Fanuc KAREL source: KD00028.KL

PROGRAM KD00028
%NOLOCKGROUP
VAR
  I: INTEGER
  J: INTEGER
  B: BOOLEAN
  R: REAL
  S: STRING[80]
BEGIN
  CONDITION[1]:
  WHEN SEMAPHORE[1] DO
    I = 1
  ENDCONDITION
END KD00028
